Fanuc KAREL source: kt00034.KL

-- PROVISIONAL review KL for V1013-1; original PC SHA256 365796e7cd78e67c99b01ca669d740d9f4b1111151055f9587d6360d3ec13897
-- Incomplete behavior may be omitted. Consult companion uncertainty JSON. Do not deploy.
PROGRAM KT00034
%NOLOCKGROUP
VAR
  I1 : INTEGER
  I2 : INTEGER
  OUT : REAL
BEGIN
  -- UNRESOLVED_PC offsets 5-16; opcodes 2E,23
  -- UNRESOLVED_PC offsets 21-32; opcodes 2E,23
  -- UNRESOLVED_PC offsets 37-48; opcodes 2E,23
  -- UNRESOLVED_PC offsets 53-64; opcodes 2E,23
  -- UNRESOLVED_PC offsets 69-89; opcodes 21,21,53,64,23
  -- UNRESOLVED_PC offsets 94-98; opcodes 7F
END KT00034
